SUBAPPLICATION GreenWhiteBackground4_AXC (* Hintergrundfarbe (TRUE -> Grün, FALSE -> Weiß) für 4 Objekte (AX-Adapter) (Kompakt) *)
  (* Standard: 61499-2 *)
  (* Version 1.0, 2026-07-21, franz, Meisterschulen am Ostbahnhof *)
  PACKAGE MyLib::sys;
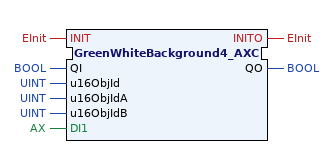
  EVENT_INPUT
    INIT : EInit; (* Initialization Request *)
  END_EVENT
  EVENT_OUTPUT
    INITO : EInit; (* Initialization Confirm *)
  END_EVENT
  VAR_INPUT
    QI : BOOL := TRUE; (* Quality Input - TRUE to enable service *)
    u16ObjId : UINT;
    u16ObjIdA : UINT;
    u16ObjIdB : UINT;
  END_VAR
  VAR_OUTPUT
    QO : BOOL; (* Quality Output - TRUE if service executed successfully *)
  END_VAR
  SOCKETS
    DI1 : adapter::types::unidirectional::AX;
  END_SOCKETS
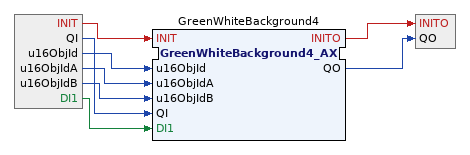
  SUBAPPS
    GreenWhiteBackground4 : MyLib::sys::GreenWhiteBackground4_AX;
  END_SUBAPPS
  EVENT_CONNECTIONS
    INIT TO GreenWhiteBackground4.INIT;
    GreenWhiteBackground4.INITO TO INITO;
  END_CONNECTIONS
  DATA_CONNECTIONS
    u16ObjId TO GreenWhiteBackground4.u16ObjId;
    u16ObjIdA TO GreenWhiteBackground4.u16ObjIdA;
    u16ObjIdB TO GreenWhiteBackground4.u16ObjIdB;
    QI TO GreenWhiteBackground4.QI;
    GreenWhiteBackground4.QO TO QO;
  END_CONNECTIONS
  ADAPTER_CONNECTIONS
    DI1 TO GreenWhiteBackground4.DI1;
  END_CONNECTIONS
END_SUBAPPLICATION
